// TIA Portal V20 export
// export: Created 2026-10-19T18:06:48.2526992Z, ExportSetting WithDefaults, DisplayName Totally Integrated Automation Portal, DisplayVersion V20 Update 6, DisplayName TIA Portal Openness, DisplayVersion V20 Update 6, DisplayName TIA Portal Version Control Interface, DisplayVersion V20 Update 6, DisplayName SINAMICS Startdrive Advanced, DisplayVersion V20 SP1, DisplayName SINAMICS Startdrive G130, G150, S120, S150, SINAMICS MV, G220, S200, S210, DisplayVersion V20 SP1, DisplayName SINAMICS Startdrive G110M, G120, G120C, G120D, G120P, G115D, DisplayVersion V20 SP1, DisplayName STEP 7 Professional, DisplayVersion V20 Update 6, DisplayName STEP 7 Safety, DisplayVersion V20 Update 2, DisplayName WinCC Basic/Comfort/Advanced, DisplayVersion V20 Update 6, DisplayName WinCC Unified, DisplayVersion V20 Update 6
DATA_BLOCK "SAI_IND_CalFree_DB"   // DB112
VERSION : 0.1
// stored: AutoNumber true, DBAccessibleFromOPCUA true, DBAccessibleFromWebserver true, InstanceOfName SAI_IND_CalFree, InstanceOfType FB
"SAI_IND_CalFree"
   // VAR_INPUT
   //    ID : HW_IO;
   // END_VAR
   // VAR_OUTPUT
   //    Process : Bool;
   //    Done : Bool;
   //    Error : Bool;
   // END_VAR
   // VAR_IN_OUT
   //    RatedCapacity : Real;
   //    Unit : SInt;
   //    RatedOutput : Real;
   //    Start : Bool;
   // END_VAR
   // VAR
   //    Activate : Bool;
   //    Status_RECORD : Int;
   //    CalFree_RECORD : Int;
   //    AdjustStep : SInt;
   //    Check01 : Bool;
   //    Check02 : Bool;
   //    WRREC_CalFree { S7_SetPoint := 'True'} : WRREC;
   //    Static01 : Bool;
   //    RDREC_Status { S7_SetPoint := 'True'} : RDREC;
   // END_VAR
BEGIN
END_DATA_BLOCK
